{attribute 'no_assign'}
FUNCTION_BLOCK FB_DO_WTURBINE_LD0_WPPD1_DevSt_st EXTENDS FB_AcsiCommonDataClass
VAR_INPUT
	stVal: FB_AcsiDATypeDevSt := (Fc:=ACSI_FC_ST, TrgOp:=ACSI_TrgOp_dchg OR ACSI_TrgOp_dupd, bLinkResult:=THIS^.AddDataToContainer(ipData:=stVal));
	q: FB_AcsiDATypeQuality := (Fc:=ACSI_FC_ST, TrgOp:=ACSI_TrgOp_qchg, bLinkResult:=THIS^.AddDataToContainer(ipData:=q));
	t: FB_AcsiDATypeTimeStamp := (Fc:=ACSI_FC_ST, bLinkResult:=THIS^.AddDataToContainer(ipData:=t));
END_VAR
VAR
END_VAR

END_FUNCTION_BLOCK

(* stored: Version 1.1.0.1
   POU FB_DO_WTURBINE_LD0_WPPD1_DevSt_st: Id {b2b1ac4b-9e11-4552-a872-2c16cc73fbaf}, SpecialFunc None *)
